(* IEC 61131-3 sources: trust-platform/examples/control/02-derivative-action-and-dynamic-response/19-poles-zeros-and-response/src, 2 files *)

(* ---- Main.st ---- *)
USING Control;

(* Pole of the first-order lag τ·dx/dt + x = K·u: the root of τs + 1 = 0. *)
FUNCTION FirstOrderPole : LREAL
VAR_INPUT
    TimeConstantS : LREAL;
END_VAR
FirstOrderPole := LREAL#-1.0 / TimeConstantS;
END_FUNCTION

(* Natural response of a real pole p: a deviation decays, or grows, as e^(p·t). *)
FUNCTION RealPoleResponse : LREAL
VAR_INPUT
    Pole : LREAL;
    Seconds : LREAL;
END_VAR
RealPoleResponse := EXP(Pole * Seconds);
END_FUNCTION

(* Poles of the shaft under P control, J·s² + B·s + Kp = 0: s = σ ± jω with σ = −B/(2J) and ω = √(Kp/J − σ²),
   a complex pair while Kp/J > σ². *)
FUNCTION ShaftPoleRealPart : LREAL
VAR_INPUT
    Inertia : LREAL;
    Friction : LREAL;
END_VAR
ShaftPoleRealPart := -Friction / (LREAL#2.0 * Inertia);
END_FUNCTION

FUNCTION ShaftPoleImaginaryPart : LREAL
VAR_INPUT
    Inertia : LREAL;
    Friction : LREAL;
    ProportionalGain : LREAL;
END_VAR
ShaftPoleImaginaryPart := SQRT(ProportionalGain / Inertia - (Friction / (LREAL#2.0 * Inertia)) ** LREAL#2.0);
END_FUNCTION

(* Unit-step response of a system with unit steady gain and the complex poles σ ± jω:
   1 − e^(σ·t)·(cos(ω·t) − (σ/ω)·sin(ω·t)). *)
FUNCTION ComplexPoleStep : LREAL
VAR_INPUT
    Sigma : LREAL;
    Omega : LREAL;
    Seconds : LREAL;
END_VAR
ComplexPoleStep := LREAL#1.0 - EXP(Sigma * Seconds) * (COS(Omega * Seconds) - Sigma / Omega * SIN(Omega * Seconds));
END_FUNCTION

PROGRAM Main
VAR
    (* The heater of Lessons 12–30 in open loop: G(s) = 0.2/(5s + 1) with the pole −0.2 s⁻¹. It rests at 36 °C
       with 80 %; the experiment returns it to 75 %, the command for 35 °C. *)
    TemperatureC : LREAL := 36.0;
    HeaterPowerPct : LREAL := 80.0;
    HeaterTimeConstantS : LREAL := 5.0;
    HeaterPole : LREAL := 0.0;
    HeaterPoleResponseC : LREAL := 36.0;
    (* The shaft of Lesson 34 under P control, Kp = 4 N·m/rad: Θ/R = 4/(s² + s + 4) with the poles −0.5 ± j1.936. *)
    Controller : Control.PID;
    Parameters : Control.PIDParameters := (
        ProportionalGain := LREAL#4.0,
        IntegralGain := LREAL#0.0,
        DerivativeGain := LREAL#0.0,
        ProportionalSetpointWeight := LREAL#1.0,
        DerivativeSetpointWeight := LREAL#0.0,
        Bias := LREAL#0.0,
        OutputMinimum := LREAL#-20.0,
        OutputMaximum := LREAL#20.0,
        RateMinimum := LREAL#-10000.0,
        RateMaximum := LREAL#10000.0,
        TrackingTime := LREAL#1.0,
        AntiWindup := PIDAntiWindup#BackCalculation
    );
    State : Control.PIDInitialState;
    Input : Control.PIDInput;
    Initialized : BOOL := FALSE;
    SetpointRad : LREAL := 0.0;
    AngleRad : LREAL := 0.0;
    VelocityRadS : LREAL := 0.0;
    TorqueNm : LREAL := 0.0;
    InertiaKgM2 : LREAL := 1.0;
    FrictionNmsRad : LREAL := 1.0;
    ShaftSigma : LREAL := 0.0;
    ShaftOmega : LREAL := 0.0;
    ShaftPoleResponseRad : LREAL := 0.0;
    (* Control Studio's project experiment starts both responses at once. *)
    ExperimentEnabled : BOOL := FALSE;
    ExperimentWasEnabled : BOOL := FALSE;
    Active : BOOL := FALSE;
    ElapsedS : LREAL := 0.0;
END_VAR

IF ExperimentEnabled AND NOT ExperimentWasEnabled THEN
    Active := TRUE;
    ElapsedS := LREAL#0.0;
ELSIF NOT ExperimentEnabled THEN
    Active := FALSE;
END_IF;
ExperimentWasEnabled := ExperimentEnabled;

IF Active THEN
    HeaterPowerPct := LREAL#75.0;
    SetpointRad := LREAL#1.0;
ELSE
    HeaterPowerPct := LREAL#80.0;
    SetpointRad := LREAL#0.0;
END_IF;

Controller.Configure(Parameters := Parameters);
IF NOT Initialized THEN
    State.Setpoint := SetpointRad;
    State.ProcessValue := AngleRad;
    Controller.Initialize(State := State);
    Initialized := TRUE;
END_IF;
Input.Mode := PIDMode#Auto;
Input.CycleTime := LREAL#0.02;
Input.Setpoint := SetpointRad;
Input.ProcessValue := AngleRad;
TorqueNm := Controller.Update(Input := Input);

(* Responses read from the poles, timed from the experiment's start. The heater's command arrives 1 s later. *)
HeaterPole := FirstOrderPole(TimeConstantS := HeaterTimeConstantS);
ShaftSigma := ShaftPoleRealPart(Inertia := InertiaKgM2, Friction := FrictionNmsRad);
ShaftOmega := ShaftPoleImaginaryPart(Inertia := InertiaKgM2, Friction := FrictionNmsRad,
    ProportionalGain := Parameters.ProportionalGain);
IF Active AND ElapsedS >= LREAL#1.0 THEN
    HeaterPoleResponseC := LREAL#35.0 + RealPoleResponse(Pole := HeaterPole, Seconds := ElapsedS - LREAL#1.0);
ELSE
    HeaterPoleResponseC := LREAL#36.0;
END_IF;
IF Active THEN
    ShaftPoleResponseRad := ComplexPoleStep(Sigma := ShaftSigma, Omega := ShaftOmega, Seconds := ElapsedS);
    ElapsedS := ElapsedS + LREAL#0.02;
ELSE
    ShaftPoleResponseRad := LREAL#0.0;
END_IF;
END_PROGRAM

CONFIGURATION Config
RESOURCE Res ON PLC
    TASK MainTask(INTERVAL := T#20ms, PRIORITY := 1);
    PROGRAM P1 WITH MainTask : Main;
END_RESOURCE
VAR_CONFIG
    P1.HeaterPowerPct AT %QL0 : LREAL;
    P1.TorqueNm AT %QL8 : LREAL;
    P1.TemperatureC AT %IL0 : LREAL;
    P1.AngleRad AT %IL8 : LREAL;
    P1.VelocityRadS AT %IL16 : LREAL;
    P1.SetpointRad AT %ML0 : LREAL;
    P1.HeaterPoleResponseC AT %ML8 : LREAL;
    P1.ShaftPoleResponseRad AT %ML16 : LREAL;
    P1.ExperimentEnabled AT %MX24.0 : BOOL;
    P1.Active AT %MX24.1 : BOOL;
END_VAR
END_CONFIGURATION

(* ---- tests.st ---- *)
(* @trustlsp:runtime-ignore — run these assertions with trust-dev test;
   they are not scheduled PLC instances in the lesson simulator. *)

TEST_PROGRAM TheHeaterPole
(* 5s + 1 = 0 at s = −0.2 s⁻¹: a 1 °C deviation decays to e^(−1) = 0.368 °C in 5 s. *)
ASSERT_NEAR(EXPECTED := LREAL#-0.2, ACTUAL := FirstOrderPole(TimeConstantS := LREAL#5.0), DELTA := LREAL#1.0e-12);
ASSERT_NEAR(EXPECTED := LREAL#0.36788,
    ACTUAL := RealPoleResponse(Pole := FirstOrderPole(TimeConstantS := LREAL#5.0), Seconds := LREAL#5.0), DELTA := LREAL#1.0e-5);
END_TEST_PROGRAM

TEST_PROGRAM TheShaftPoles
VAR
    Sigma : LREAL;
    Omega : LREAL;
END_VAR
(* s² + s + 4 = 0 at s = −0.5 ± j1.9365: a swing every 2π/ω = 3.245 s; the first peak at π/ω = 1.622 s reaches
   1 + e^(−0.5·1.622) = 1.444 rad. *)
Sigma := ShaftPoleRealPart(Inertia := LREAL#1.0, Friction := LREAL#1.0);
Omega := ShaftPoleImaginaryPart(Inertia := LREAL#1.0, Friction := LREAL#1.0, ProportionalGain := LREAL#4.0);
ASSERT_NEAR(EXPECTED := LREAL#-0.5, ACTUAL := Sigma, DELTA := LREAL#1.0e-12);
ASSERT_NEAR(EXPECTED := LREAL#1.93649, ACTUAL := Omega, DELTA := LREAL#1.0e-5);
ASSERT_NEAR(EXPECTED := LREAL#3.24462, ACTUAL := LREAL#2.0 * LREAL#3.14159265358979 / Omega, DELTA := LREAL#1.0e-5);
ASSERT_NEAR(EXPECTED := LREAL#1.44434,
    ACTUAL := ComplexPoleStep(Sigma := Sigma, Omega := Omega, Seconds := LREAL#3.14159265358979 / Omega), DELTA := LREAL#1.0e-5);
(* Kp = 16: s = −0.5 ± j3.969, a swing every 1.583 s inside the same envelope e^(−0.5t). *)
ASSERT_NEAR(EXPECTED := LREAL#3.96863,
    ACTUAL := ShaftPoleImaginaryPart(Inertia := LREAL#1.0, Friction := LREAL#1.0, ProportionalGain := LREAL#16.0), DELTA := LREAL#1.0e-5);
END_TEST_PROGRAM

TEST_PROGRAM ThePiLoopPolesAndZeros
VAR
    S : LREAL;
END_VAR
(* PI on the heater without delay, C = 2.5 + 0.5/s: 1 + CG = 0 gives 5s² + 1.5s + 0.1 = 0, the poles −0.1 and −0.2.
   The setpoint numerator 0.5s + 0.1 has its zero at −0.2; the disturbance numerator 0.2s at 0. *)
S := LREAL#-0.1;
ASSERT_NEAR(EXPECTED := LREAL#0.0, ACTUAL := LREAL#5.0 * S * S + LREAL#1.5 * S + LREAL#0.1, DELTA := LREAL#1.0e-12);
S := LREAL#-0.2;
ASSERT_NEAR(EXPECTED := LREAL#0.0, ACTUAL := LREAL#5.0 * S * S + LREAL#1.5 * S + LREAL#0.1, DELTA := LREAL#1.0e-12);
ASSERT_NEAR(EXPECTED := LREAL#0.0, ACTUAL := LREAL#0.5 * S + LREAL#0.1, DELTA := LREAL#1.0e-12);
(* A 1 % disturbance step: x(t) = 0.4·(e^(−0.1t) − e^(−0.2t)) °C, largest at t = ln 2/0.1 = 6.93 s with 0.1 °C. *)
ASSERT_NEAR(EXPECTED := LREAL#0.1,
    ACTUAL := LREAL#0.4 * (RealPoleResponse(Pole := LREAL#-0.1, Seconds := LN(LREAL#2.0) / LREAL#0.1)
        - RealPoleResponse(Pole := LREAL#-0.2, Seconds := LN(LREAL#2.0) / LREAL#0.1)), DELTA := LREAL#1.0e-12);
END_TEST_PROGRAM
